(* IEC 61131-3 sources: plc-vscode/tests/st/all/rusty/tests/lit/single/address, 8 files *)

(* ---- fn_local_at_round_trip.st ---- *)
// RUN: (%COMPILE %s && %RUN) | %CHECK %s
// Probe for #1737 follow-up: a FUNCTION-scoped VAR with `AT %M...` should bind its alias
// pointer to the synthesised backing global on entry, so the write below ends up at the
// same hardware slot a VAR_GLOBAL alias would observe.

VAR_GLOBAL
    g AT %MX1.2.3.4 : BYTE;
END_VAR

FUNCTION writer : DINT
VAR
    local AT %MX1.2.3.4 : BYTE;
END_VAR
    local := 7;
    writer := DINT#0;
END_FUNCTION

FUNCTION main : DINT
    writer();
    // CHECK: 7
    printf('%d$N', g);
END_FUNCTION

(* ---- hardware_reference_used.st ---- *)
// RUN: (%COMPILE %s && %RUN) | %CHECK %s
VAR_GLOBAL
    a AT %IX1.2.1 : BOOL;
    b AT %QX1.2.2 : BOOL;
    c AT %ID1.2.3 : DWORD;
    d AT %ID1.2.4 : DWORD;
END_VAR

FUNCTION main : DINT
    a := TRUE;
    printf('%u$N', a); //CHECK: 1
    b := TRUE;
    printf('%u$N', b); //CHECK: 1
    c := 1337;
    printf('%d$N', c); //CHECK: 1337
    d := 98765;
    printf('%d$N', d); //CHECK: 98765
END_FUNCTION

(* ---- reference_in_body.st ---- *)
// RUN: (%COMPILE %s && %RUN) | %CHECK %s
VAR_GLOBAL
    a AT %IX1.2.1 : BOOL;
    b AT %QX1.2.2 : BOOL;
    c AT %ID1.2.3 : DWORD;
    d AT %ID1.2.4 : DWORD;
END_VAR

FUNCTION main : DINT
    %IX1.2.1 := TRUE;
    printf('%u$N', a); //CHECK: 1
    b := TRUE;
    printf('%u$N', %QX1.2.2); //CHECK: 1
    %IX1.2.3 := 1337;
    printf('%d$N', c); //CHECK: 1337
    d := 98765;
    printf('%d$N', %QX1.2.4); //CHECK: 98765
END_FUNCTION

(* ---- method_var_at_round_trip.st ---- *)
// RUN: (%COMPILE %s && %RUN) | %CHECK %s
// #1737 coverage: a METHOD-scoped VAR with `AT %M...` should alias-bind on method
// entry and round-trip a write to the backing hardware slot.

VAR_GLOBAL
    g AT %MX3.4.5.6 : BYTE;
END_VAR

FUNCTION_BLOCK probeFb
    METHOD writer
    VAR
        local AT %MX3.4.5.6 : BYTE;
    END_VAR
        local := 17;
    END_METHOD
END_FUNCTION_BLOCK

PROGRAM mainProg
VAR
    p : probeFb;
END_VAR
    p.writer();
END_PROGRAM

FUNCTION main : DINT
    mainProg();
    // CHECK: 17
    printf('%d$N', g);
END_FUNCTION

(* ---- method_var_temp_at_round_trip.st ---- *)
// RUN: (%COMPILE %s && %RUN) | %CHECK %s
// #1737 coverage: a METHOD-scoped VAR_TEMP with `AT %M...` (temporary, per-call) should
// alias-bind on entry and round-trip a write to the backing hardware slot.

VAR_GLOBAL
    g AT %MX4.5.6.7 : BYTE;
END_VAR

FUNCTION_BLOCK probeFb
    METHOD writer
    VAR_TEMP
        local AT %MX4.5.6.7 : BYTE;
    END_VAR
        local := 23;
    END_METHOD
END_FUNCTION_BLOCK

PROGRAM mainProg
VAR
    p : probeFb;
END_VAR
    p.writer();
END_PROGRAM

FUNCTION main : DINT
    mainProg();
    // CHECK: 23
    printf('%d$N', g);
END_FUNCTION

(* ---- var_global_and_fb_share_hw_address.st ---- *)
// RUN: (%COMPILE %s && %RUN) | %CHECK %s
// Issue #1736: a complete hardware address (AT %MX1.2.3.4) on a POU-scoped variable used to be
// silently dropped at codegen — the FB field stayed null and the first access SIGSEGV'd at
// runtime. The preprocessor now synthesises the backing __M_1_2_3_4 global and the existing
// alias-pointer lowering binds the FB field in the per-instance ctor. The VAR_GLOBAL `slot`
// and the FB `shadow` must end up bound to the *same* `__M_1_2_3_4` slot.

VAR_GLOBAL
    slot AT %MX1.2.3.4 : BYTE;
END_VAR

FUNCTION_BLOCK probe
VAR_INPUT
    shadow AT %MX1.2.3.4 : BYTE;
END_VAR
    shadow := 42;
END_FUNCTION_BLOCK

PROGRAM mainProg
VAR
    p : probe;
END_VAR
    p();
    // CHECK: 42
    printf('%d$N', slot);
END_PROGRAM

FUNCTION main : DINT
    mainProg();
END_FUNCTION

(* ---- alias_hardware_roundtrip.st ---- *)
// RUN: (%COMPILE %s && %RUN) | %CHECK %s
VAR_GLOBAL
    alias AT %IX1.1 : BOOL;
END_VAR

PROGRAM prog
VAR
    tmp : BOOL;
END_VAR
    // CHECK: 1
    alias := TRUE;
    tmp := %IX1.1;
    printf('%u$N', tmp);

    // CHECK: 0
    %IX1.1 := FALSE;
    tmp := alias;
    printf('%u$N', tmp);
END_PROGRAM

FUNCTION main : DINT
    prog();
END_FUNCTION

(* ---- program_local_at_round_trip.st ---- *)
// RUN: (%COMPILE %s && %RUN) | %CHECK %s
// #1737 coverage: a PROGRAM-scoped VAR with `AT %M...` should bind its alias on the
// per-instance ctor, so the write below ends up at the same hardware slot a
// VAR_GLOBAL alias at the same address observes.

VAR_GLOBAL
    g AT %MX2.3.4.5 : BYTE;
END_VAR

PROGRAM probeProg
VAR
    local AT %MX2.3.4.5 : BYTE;
END_VAR
    local := 11;
END_PROGRAM

FUNCTION main : DINT
    probeProg();
    // CHECK: 11
    printf('%d$N', g);
END_FUNCTION
